(* IEC 61131-3 sources: daoli-st-library/DL_Base (part 21) *)

(* ---- FC_DL_BitArrayExtract.st ---- *)
(*==============================================================================
 * 组件名称 (Component)  : FC_DL_BitArrayExtract
 * 所属子库 (Sublibrary) : DL_Base
 * 归属目录 (Directory)  : C:\Library\DL_Base
 * 当前版本 (Version)    : 1.0.0
 * 组件分类 (Category)   : 函数（FUNCTION）· 纯函数 · 跨字位流窗口提取
 * 兼容性   (Platform)   : CODESYS 3.5 / TwinCAT 3 / 汇川 InoProShop / 施耐德
 *                         Machine Expert；仅用 Standard.library 的 SHL / SHR /
 *                         AND / OR 与显式类型转换，无厂商位访问方言，无实例依赖
 * 功能一句话 (Summary)  : 从 DWORD 数组构成的连续位流中按「起始位 + 位宽」取出
 *                         位窗口并右对齐输出，同时给出本次生效掩码。
 * 功能描述 (Function)   : 第 1 个数组元素承载位 0 到 31，第 2 个承载位 32 到 63，
 *                         依此类推（LSB 起）。调用方给出起始位与位宽，本件负责
 *                         跨字拼接、右移对齐、掩码构造与三类边界拦截。
 *                         典型现场用途：64 位设备状态字经两个保持寄存器上传后的
 *                         字段解码、凸轮表位图跨 4 个双字存放时的段取出、
 *                         远程 IO 位图跨字存放时的报警位段读取。
 * 与既有件边界 (Boundary): FC_DL_BitGet 取单字内单个位；FC_DL_BitFieldExtract 取
 *                         单字内 1 到 32 位段；FB_DL_UnpackWordToBits 把单字拆成
 *                         16 个固定位。三者都只作用于一个 32 位字。本件是「跨字
 *                         位流窗口」，位窗可跨 2 个双字、宽度可达 64 位，四者职责
 *                         互斥，不复用也不替代其中任何一件。
 * 设计要点 (Key notes)  : ① 闸门顺序固定为「字数 → 偏移 → 宽度 → 越界截断」，
 *                           任一闸门拦下即预置输出后返回，绝不让非法移位量进入
 *                           SHL / SHR（越界移位在部分编译器属未定义行为）；
 *                         ② 宽度 64 走满 1 常量分支，禁止 SHL(x, 64)；
 *                         ③ 截断只报事件不返回空值：现场宁可读到半段有效位，
 *                           由调用方依据 bValid 与 nActualW 自行判断完整度；
 *                         ④ 纯函数：无内部状态、无跨周期残留，同入参同结果。
 * 开源溯源 (Origin)     : 来源标签 lgf-bitlogic。LGF（Libre Graphical Framework）
 *                         为免费闭源发布的公开函数库手册，本件仅借鉴其位逻辑组
 *                         「单点 → 单段 → 批量段」的分层分类，以及「源 / 起位 /
 *                         位宽」三段参数域的组织方式；许可证按其发布方条款仅作
 *                         分类参考，本件零代码行、零注释、零数据结构引用，
 *                         属 clean-room 独立实现，不构成衍生作品。
 * 码位说明 (Codes)      : 本件独占信息级码段 16#0001_0125 到 16#0001_0127，纯函数
 *                         无锁存面故不占故障级码；三段与全库已占码求差为空，
 *                         不与 DL_MathData 的 0101 到 0124 任何一件重叠。
 *                         0125 偏移越界 ｜ 0126 宽度越界 ｜ 0127 跨字截断。
 * 依赖说明 (Depends)    : 无 DL_ 内部依赖；仅 Standard.library 的 SHL / SHR /
 *                         DWORD_TO_LWORD / INT_TO_DINT / INT_TO_UDINT。
 * 契约前置条件 (Contract): 入参为数组形参，函数内无法探测数组实际长度，故
 *                         「nSourceCount 不得大于调用方实际数组长度」由调用方负责。
 *                         这是本库唯一允许的契约式前置条件，调用方须在组态时保证。
 * 红线自检 (Redline)    : 零全局变量表依赖 ｜ 零外部变量声明 ｜ 零物理地址
 *                         纯 IEC 61131-3 ｜ 无除法故无除零面 ｜ 全变量双语同行注释
 *                         状态机 N/A（纯函数）｜ 无定时器实例
 * 修订历史 (Revision)   : 2026-11-15  v1.0.0  首版入库（Round 12 · 跨字位段族）
 *============================================================================*)

(*==============================================================================
 * 位流几何示意 (Bit stream geometry)：
 *   auSource[1] 承载位 0 到 31，auSource[2] 承载位 32 到 63，位号自低向高
 *   以 auSource[1] = 16#1234_5678、auSource[2] = 16#9ABC_DEF0 为例：
 *     拼接后的 64 位窗口为 16#9ABCDEF0_12345678
 *     起始位 28、位宽 8 取出的是位 28 到 35：低位 4 位来自第 1 字最高半字节，
 *     高位 4 位来自第 2 字最低半字节，右对齐结果为 16#01
 *     起始位 20、位宽 16 取出的位 20 到 35，右对齐结果为 16#0123
 *============================================================================*)

(*==============================================================================
 * 逐调用推演 (Call trace)：
 *   调用 1  两字、起始 28、位宽 8
 *     字数为 2，总位数 64；偏移 28 小于 64 通过；宽度 8 在 1 到 64 内通过
 *     28 加 8 等于 36 不超过 64，不截断
 *     低字下标 1，字内移位 28，28 加 8 大于 32 且 1 小于 2，高字下标 2
 *     拼接右移 28 位后取低 8 位，得 16#01，掩码 16#FF，有效
 *   调用 2  同上两字、起始 28、位宽 40
 *     28 加 40 等于 68 超过 32 位窗口可覆盖范围，宽度截为 4，事件码 0127
 *     结果只含 4 位可用值，bValid 为假，但值仍可读
 *   调用 3  起始 32、字数 1
 *     总位数 32，偏移不小于总位数，早退，事件码 0125，输出全零
 *============================================================================*)

(*==============================================================================
 * 调用示例 (Instance guide)：
 *   bOk := FC_DL_BitArrayExtract(
 *              auSource     := aStatusWords,
 *              nSourceCount := 2,
 *              nOffset      := 28,
 *              nWidth       := 8,
 *              uField       => uFieldOut,
 *              nActualW     => nWidthUsed);
 *   提示：uField 已右对齐，比较时应与右对齐期望值比较；判定完整度请看 bValid。
 *============================================================================*)

FUNCTION FC_DL_BitArrayExtract : BOOL
VAR_IN_OUT
    auSource     : ARRAY[1..8] OF DWORD;  // 源位流数组，第 1 元素为位 0 到 31，第 2 元素为位 32 到 63 [位串] / Source bit stream, element 1 holds bits 0 to 31
END_VAR
VAR_INPUT
    nSourceCount : INT := 1;              // 源有效字数 [个]，域 1 到 8，越界钳位 / Effective source word count, 1 to 8, clamped
    nOffset      : INT := 0;              // 位窗口起始位 [bit]，0 起，域 0 到 32 乘字数减 1 / Window start bit, zero based
    nWidth       : INT := 1;              // 位窗口宽度 [bit]，域 1 到 64 / Window width, 1 to 64
END_VAR
VAR_OUTPUT
    uField       : LWORD;                 // 右对齐提取结果，bit0 起连续 nActualW 位有效 [位串] / Extracted field, right aligned
    uMask        : LWORD;                 // 本次实际生效掩码，已右对齐，可直接与结果位与 [位串] / Effective right aligned mask
    nActualW     : INT;                   // 实际生效宽度，越界截断后的值 [bit] / Effective width after truncation
    uErrorId     : UDINT;                 // 事件码，0 表示无事件 / Event code, zero means none
    bValid       : BOOL;                  // 入参域全合法为真，发生截断或越界为假（截断时结果仍可用） / Inputs legal, false when truncated
END_VAR
VAR
    nTotalBits   : DINT;                  // 位流总位数，等于字数乘 32，DINT 中间量防 INT 溢出 [bit] / Total bit count, DINT to avoid overflow
    nIdxLo       : INT;                   // 低字下标，1 起 [索引] / Low word index, one based
    nIdxHi       : INT;                   // 高字下标，1 起，不跨字时置 0 [索引] / High word index, zero when not straddling
    uWide        : LWORD;                 // 两字拼接的 64 位窗口值 [位串] / Stitched 64 bit window
    uLo          : DWORD;                 // 低字快照 [位串] / Low word snapshot
    uHi          : DWORD;                 // 高字快照，不跨字时为 0 [位串] / High word snapshot, zero when absent
    nShift       : INT;                   // 字内移位量，等于偏移对 32 取模 [bit] / Intra word shift amount
END_VAR
VAR CONSTANT
    DL_SRC_MAX    : INT := 8;                          // 源字数上限 [个] / Source word count limit
    DL_BIT_MAX64  : INT := 64;                         // 位窗宽度上限 [bit] / Window width limit
    DL_BIT_MAX32  : INT := 32;                         // 单字位宽 [bit] / Bits per word
    DL_MASK64_ALL : LWORD := 16#FFFF_FFFF_FFFF_FFFF;   // 满宽掩码常量，64 宽分支专用 [位串] / All ones mask for the 64 bit branch
    DL_GUARD_MAX  : DINT := 64;                        // 循环守卫上限，本件直线实现无循环体，按组件族口径保留 [次] / Loop guard limit kept by family convention, no loop here
END_VAR

(*------------------------------------------------------------------------------
 * 段 1｜输出预置：任何异常路径下输出必须确定
 *      Pre-set outputs so that every path is deterministic
 *-----------------------------------------------------------------------------*)
FC_DL_BitArrayExtract := FALSE;
uField                := 16#0000_0000_0000_0000;
uMask                 := 16#0000_0000_0000_0000;
nActualW              := 0;
uErrorId              := 16#0000_0000;
bValid                := FALSE;

(*------------------------------------------------------------------------------
 * 段 2｜源字数钳位（边界 B1）：先夹到 1 到 8，再算总位数
 *      Clamp the word count first, then derive the total bit count
 *-----------------------------------------------------------------------------*)
IF nSourceCount < 1 THEN
    nSourceCount := 1;
ELSIF nSourceCount > DL_SRC_MAX THEN
    nSourceCount := DL_SRC_MAX;
END_IF
nTotalBits := INT_TO_DINT(nSourceCount) * INT_TO_DINT(DL_BIT_MAX32);

(*------------------------------------------------------------------------------
 * 段 3｜偏移闸门（边界 B2）：负偏移与落空偏移一律早退
 *      Offset gate: negative or beyond the stream end exits early
 *-----------------------------------------------------------------------------*)
IF (nOffset < 0) OR (INT_TO_DINT(nOffset) >= nTotalBits) THEN
    uErrorId := 16#0001_0125;   // 偏移越界，输出保持全零
    RETURN;
END_IF

(*------------------------------------------------------------------------------
 * 段 4｜宽度闸门（边界 B3）：宽度须落在 1 到 64 闭区间
 *      Width gate: the window width must be within one to sixty four
 *-----------------------------------------------------------------------------*)
IF (nWidth < 1) OR (nWidth > DL_BIT_MAX64) THEN
    uErrorId := 16#0001_0126;   // 宽度越界，输出保持全零
    RETURN;
END_IF

(*------------------------------------------------------------------------------
 * 段 5｜越界截断（边界 B4）：按位流末端截断，仍继续计算可用低位
 *      Truncation at the stream end: the usable low bits are still produced
 *      工程取舍：不返空值，现场宁可读半段，完整度交给 bValid 判断
 *-----------------------------------------------------------------------------*)
IF (INT_TO_DINT(nOffset) + INT_TO_DINT(nWidth)) > nTotalBits THEN
    nWidth   := DINT_TO_INT(nTotalBits - INT_TO_DINT(nOffset));
    uErrorId := 16#0001_0127;
    bValid   := FALSE;
END_IF

(*------------------------------------------------------------------------------
 * 段 6｜定位（边界 B5）：求低字下标与字内移位量，判断是否跨字
 *      Locate the low word and the intra word shift, decide straddling
 *      nShift 由取模保证 0 到 31，负移位量不可能出现
 *-----------------------------------------------------------------------------*)
nIdxLo := nOffset / DL_BIT_MAX32 + 1;
nShift := nOffset MOD DL_BIT_MAX32;
nIdxHi := 0;
IF ((nShift + nWidth) > DL_BIT_MAX32) AND (nIdxLo < nSourceCount) THEN
    nIdxHi := nIdxLo + 1;
END_IF

(*------------------------------------------------------------------------------
 * 段 7｜双字窗口深度校验（边界 B6）：位窗跨越第三个字时按双字窗口截断
 *      Third word guard: a window reaching the next word is truncated here
 *      原因：移位中间量为 64 位，起点非零时最多只能覆盖到第二个字末尾，
 *      若不截断则高位会静默读成零；此处显式截断并报事件，杜绝静默错值
 *-----------------------------------------------------------------------------*)
IF (nShift + nWidth) > DL_BIT_MAX64 THEN
    nWidth   := DL_BIT_MAX64 - nShift;
    uErrorId := 16#0001_0127;
    bValid   := FALSE;
END_IF

(*------------------------------------------------------------------------------
 * 段 8｜拼接（边界 B7）：先取低字，跨字时把高字左移 32 位后并入
 *      Stitch low word first, then merge the high word shifted by 32
 *      下标安全性：偏移已验证小于总位数，故低字下标不超过字数上限；
 *      高字下标仅在下标小于字数时置位，越界读取不可能发生
 *-----------------------------------------------------------------------------*)
uLo   := auSource[nIdxLo];
uHi   := 16#0000_0000;
IF nIdxHi > 0 THEN
    uHi := auSource[nIdxHi];
END_IF
uWide := DWORD_TO_LWORD(uLo);
IF nIdxHi > 0 THEN
    uWide := uWide OR SHL(DWORD_TO_LWORD(uHi), DL_BIT_MAX32);
END_IF

(*------------------------------------------------------------------------------
 * 段 9｜右对齐：整体右移字内移位量，移位量 0 到 31 必在合法域
 *      Right align by shifting the stitched window down
 *-----------------------------------------------------------------------------*)
uWide := SHR(uWide, INT_TO_UDINT(nShift));

(*------------------------------------------------------------------------------
 * 段 10｜掩码构造（边界 B8）：64 宽走满一常量分支，禁止左移 64 位
 *      Mask construction: the full width case uses the constant branch
 *-----------------------------------------------------------------------------*)
IF nWidth >= DL_BIT_MAX64 THEN
    uMask := DL_MASK64_ALL;
ELSE
    uMask := SHL(LWORD#1, INT_TO_UDINT(nWidth)) - LWORD#1;
END_IF

(*------------------------------------------------------------------------------
 * 段 11｜结果收口：掩码与窗口相与，宽度与有效位一次性定稿
 *      Close out: mask the window and publish the effective width
 *-----------------------------------------------------------------------------*)
uField   := uWide AND uMask;
nActualW := nWidth;
IF uErrorId = 16#0000_0000 THEN
    bValid                := TRUE;
    FC_DL_BitArrayExtract := TRUE;
END_IF
END_FUNCTION

(* ---- FC_DL_BitArrayRotate.st ---- *)
(*==============================================================================
 * 组件名称 (Component)  : FC_DL_BitArrayRotate
 * 所属子库 (Sublibrary) : DL_Base
 * 归属目录 (Directory)  : C:\Library\DL_Base
 * 当前版本 (Version)    : 1.0.0
 * 分类/来源标签         : 函数（FUNCTION）· 纯函数 · 跨字整串循环移位
 *                         lgf-bitlogic / bit-manipulation / cross-word
 * 兼容性   (Platform)   : CODESYS 3.5 / TwinCAT 3 / 汇川 InoProShop / 施耐德
 *                         Machine Expert；仅用 Standard.library 的 SHL / SHR /
 *                         OR / ABS 与显式类型转换，无厂商位访问方言，无实例依赖
 * 功能一句话 (Summary)  : 把 1 到 4 个 DWORD 视为一条 32 到 128 位的位串，整体
 *                         左移或右移 n 位，移出最高字的位回卷到最低字。
 * 功能描述 (Function)   : 第 1 个数组元素承载位 0 到 31，第 2 个承载位 32 到 63，
 *                         依此类推（每字内 LSB 起）。整体旋转与单字循环移位不同：
 *                         位串总宽 W 等于 32 乘有效字数，左移 s 位时目标位 i 取自
 *                         源位 (i 减 s) 对 W 取模，因此最高字移出的位回卷到第 1 字
 *                         最低位。典型现场用途：多字报警位图的时段轮转显示、
 *                         4 字 128 点位图的交接班整体顺延、循环缓冲区位索引的
 *                         整体平移、旋转编码器多字计数的位窗口对齐。
 * 与既有件边界 (Boundary): FC_DL_BitArrayExtract 是「抽」、FC_DL_BitArrayInsert 是
 *                         「插」、本件是「转」。前两件按位窗口做局部读写，本件只做
 *                         整条位串的循环平移，位序总量守恒、位宽不变。三者构成
 *                         位段族三件套，职责互斥、参数域不重叠。
 * 为什么不用标准 ROL     : IEC 的 ROL 只在单字内循环，跨字无定义；多字拼成 64 位
 *                         或 128 位中间量再移位的写法，在移位量等于位宽时属未定义
 *                         行为，且各平台对超宽中间量的支持不一致。本件按字就地
 *                         运算，移位量一律落在 1 到 31 的合法域。
 * 设计要点 (Key notes)  : ① 闸门顺序固定为「字数 → 移位归约 → 逐字合成」，字数非法
 *                           直接早退且不写目标；
 *                         ② 移位量先取绝对值再对总宽取模，永远不把原始 nShift 送进
 *                           SHL / SHR；
 *                         ③ 方向归一裁定：nShift 的符号优先于 bLeft，负值恒为右移，
 *                           非负时由 bLeft 决定左或右（详见下方方向表）；
 *                         ④ 结果先落到局部暂存数组，全部算完再整体写回，因而目标
 *                           与源同址（别名）时不会读到被覆盖的中间值；
 *                         ⑤ 纯函数：无内部状态、无跨周期残留，同入参同结果。
 *
 * 【方向归一表 / Direction normalisation table】
 *   nShift < 0            → 右移，量取绝对值，bLeft 被忽略
 *   nShift >= 0, bLeft    → 左移，量为 nShift
 *   nShift >= 0, bLeft 假 → 右移，量为 nShift
 *   左移量最终统一折算成 0 到 W 减 1 的左旋量，右移按「W 减量」等值换算
 *
 * 【验收向量 / Acceptance vectors】
 *   V1  nWords=2, aSrc=[16#8000_0001, 16#0000_0000], nShift=1, bLeft=真
 *       → aDst=[16#0000_0002, 16#0000_0001]，nEffectiveShift=1（最高位回卷第 2 字）
 *   V2  nWords=2, 同一源, nShift=1, bLeft=假
 *       → aDst=[16#4000_0000, 16#8000_0000]，nEffectiveShift=63（最低位回卷最高字）
 *   V3  V-B 边界：nWords=2, nShift=64 → 归约后 nEffectiveShift=0，输出等于输入，
 *       置 013D（整圈也是「移位量被归约」，必须有人说一声）
 *   V4  V-A 域外：nWords=0 → 返回 FALSE、021F、aDst 原样不动（不写半张图）
 *   V5  V-B 边界：nWords=9 → 钳到 4、置 013E、按 4 字旋转
 *   V6  单字：nWords=1, aSrc[1]=16#8000_0001, nShift=1, bLeft=真
 *       → aDst[1]=16#0000_0003（单字内首尾位同时回卷，验证取模路径）
 *
 * 开源溯源 (Origin)     : 来源标签 lgf-bitlogic。LGF（Libre Graphical Framework）
 *                         为免费闭源发布的公开函数库手册，本件仅借鉴其位逻辑组
 *                         「单点、单段、批量段」的分层分类，以及「源、目标、移位量」
 *                         三段参数域的组织方式；许可证按其发布方条款仅作分类参考，
 *                         本件零代码行、零注释、零数据结构引用，属 clean-room
 *                         独立实现，不构成衍生作品。
 * 码位说明 (Codes)      : 信息 16#0001_013D 移位量已归约 ｜ 16#0001_013E 字数已钳位
 *                         故障 16#0001_021F 字数非法。三段取号见本轮规格 §3.2，
 *                         与位段族既有 0125 到 0127 区间不重叠。
 * 依赖说明 (Depends)    : 无 DL_ 内部依赖；仅 Standard.library 的 SHL / SHR /
 *                         ABS 与 INT_TO_DINT / DINT_TO_INT。
 * 契约前置条件 (Contract): 入参为定长数组形参，函数内无法探测调用方数组实际长度，
 *                         故「nWords 不得大于调用方数组长度」由调用方在组态时保证。
 * 镜像量清单 (R38)      : 本件无锁存副本，边界量全部由入口标量 nWords 与 nShift
 *                         自身导出，不存在锁存量与实时量混用面。
 * 红线自检 (Redline)    : 零全局变量表依赖 ｜ 零外部变量声明 ｜ 零物理地址直写
 *                         纯 IEC 61131-3 ｜ 无除法故无除零面 ｜ 空移位量走常量分支
 *                         全变量双语同行注释 ｜ 状态机 N/A（纯函数）｜ 无定时器实例
 * 修订历史 (Revision)   : 2026-11-15  v1.0.0  首版入库（Round 13 · 泳道 B 位段族收口）
 *============================================================================*)

(*==============================================================================
 * 位串几何示意 (Bit string geometry)：
 *   两字共 64 位，位 0 到 31 在第 1 字，位 32 到 63 在第 2 字
 *   源 16#8000_0001 与 16#0000_0000 的置位点是位 0 与位 31
 *   左旋 1 位：位 0 到 1、位 31 到 32，故结果第 1 字 16#0000_0002、
 *   第 2 字 16#0000_0001，位宽守恒（仍是两个置位点）
 *   右旋 1 位：位 0 到 63、位 31 到 30，故结果第 1 字 16#4000_0000、
 *   第 2 字 16#8000_0000
 *============================================================================*)

(*==============================================================================
 * 逐调用推演 (Call trace)：
 *   调用 1  两字、左移 1
 *     字数 2 合法；总宽 64；左移量 1，对 64 取模仍为 1，k 为 0、r 为 1
 *     第 1 字取源字 1 左移 1 或源字 2 右移 31，得 16#0000_0002
 *     第 2 字取源字 2 左移 1 或源字 1 右移 31，得 16#0000_0001
 *   调用 2  两字、右移 1
 *     折算左旋量 64 减 1 等于 63，k 为 1、r 为 31
 *     r 非零，第 1 字取源字 2 左移 31 或源字 1 右移 1，得 16#4000_0000
 *   调用 3  字数 0
 *     闸门 1 拦下，返回假、码 021F，目标数组一次都没写
 *============================================================================*)

(*==============================================================================
 * 调用示例 (Instance guide)：
 *   bOk := FC_DL_BitArrayRotate(
 *              aSrc            := aAlarmMap,
 *              nWords          := 4,
 *              nShift          := 8,
 *              bLeft           := TRUE,
 *              aDst            := aAlarmMapShifted,
 *              nEffectiveShift => nUsed,
 *              uErrorId        => uCode);
 *   提示：nEffectiveShift 是归约后的左旋量，不是入参原值；要判「有没有整圈」
 *         请比对 16#0001_013D 是否出现。
 *============================================================================*)

FUNCTION FC_DL_BitArrayRotate : BOOL
VAR_INPUT
    aSrc   : ARRAY[1..4] OF DWORD;  // 源位图，第 1 元素为位 0 到 31，未用字填 0 [位串] / Source bitmap, element 1 holds bits 0 to 31, unused words zeroed
    nWords : INT;                   // 有效字数 [个]，域 1 到 4，越界按钳位规则处理 / Effective word count, 1 to 4, clamped
    nShift : INT;                   // 移位位数 [bit]，负值恒为右移，域负 32767 到 32767 / Shift amount, negative always means right
    bLeft  : BOOL;                  // 方向选择，真为左移（向高位），假为右移；nShift 为负时本引脚被忽略 / TRUE rotates left, ignored when nShift is negative
END_VAR
VAR_IN_OUT
    aDst   : ARRAY[1..4] OF DWORD;  // 目标位图，允许与源同址；失败路径不写入 [位串] / Destination bitmap, may alias the source, untouched on failure
END_VAR
VAR_OUTPUT
    nEffectiveShift : INT;          // 归一后实际左旋量 [bit]，域 0 到总宽减 1 / Effective left rotation after normalisation
    uErrorId        : UDINT;        // 事件码，0 表示无事件 / Event code, zero means none
END_VAR
VAR
    nW        : INT;                // 钳位后的有效字数 [个] / Clamped effective word count
    nWidthBit : DINT;               // 位串总宽，等于字数乘 32，DINT 中间量防溢出 [bit] / Total bit width in DINT
    nMag      : DINT;               // 移位量绝对值 [bit] / Absolute shift magnitude
    nMod      : DINT;               // 绝对值对总宽取模的结果 [bit] / Magnitude reduced modulo the width
    nLeft     : DINT;               // 折算后的左旋量 [bit]，域 0 到总宽减 1 / Normalised left rotation amount
    nWordOfs  : DINT;               // 左旋量折算的整字偏移 k [字] / Whole word offset derived from the rotation
    nBitOfs   : INT;                // 左旋量折算的字内偏移 r [bit]，域 0 到 31 / Intra word offset, 0 to 31
    bRight    : BOOL;               // 实际方向，真为右移 / Effective direction, TRUE means right
    nJ        : INT;                // 目标字下标，1 起 [索引] / Destination word index, one based
    nIdxA     : INT;                // 左移贡献源字的下标，0 起算后加 1 [索引] / Source index for the left shifted contribution
    nIdxB     : INT;                // 右移贡献源字的下标，0 起算后加 1 [索引] / Source index for the right shifted contribution
    uA        : DWORD;              // 左移贡献源字快照 [位串] / Snapshot of the left shifted source word
    uB        : DWORD;              // 右移贡献源字快照 [位串] / Snapshot of the right shifted source word
    aTmp      : ARRAY[1..4] OF DWORD;   // 结果暂存区，全部算完才写回目标，保证别名安全 [位串] / Staging buffer, written back only after the whole result is ready
END_VAR
VAR CONSTANT
    DL_BAR_MAXW  : INT := 4;    // 最大字数 [个]，与形参维度字面量一致 / Maximum word count, must match the array dimension
    DL_BAR_WBITS : INT := 32;   // 单字位宽 [bit] / Bits per word
    DL_BAR_SHMAX : DINT := 127; // 规格允许的移位量绝对值上限 [bit] / Documented shift magnitude limit
END_VAR

(*------------------------------------------------------------------------------
 * 段 1｜输出预置：任何路径下的可读输出必须确定
 *      Pre-set the readable outputs so every path is deterministic
 *      目标数组刻意不预置：失败契约要求「原样不动」，先写就破了契约
 *      The destination is deliberately left untouched, the failure contract keeps it as is
 *-----------------------------------------------------------------------------*)
FC_DL_BitArrayRotate := FALSE;
nEffectiveShift     := 0;
uErrorId            := 16#0000_0000;
nW                  := 0;
nBitOfs             := 0;
nWordOfs            := 0;
bRight              := FALSE;
nMod                := 0;
nLeft               := 0;

(*------------------------------------------------------------------------------
 * 段 2｜字数闸门（边界 B1/B2）：小于 1 属逻辑错，早退且不写目标
 *      Word count gate: below one is a logic error, exit early without writing
 *      大于 4 属契约超界，钳位后照算，现场宁可转错半张图也不要空输出
 *      Above four is a contract breach, clamped and still computed
 *-----------------------------------------------------------------------------*)
IF nWords < 1 THEN
    uErrorId := 16#0001_021F;   // 故障级：字数非法，目标数组保持原样
    RETURN;
ELSIF nWords > DL_BAR_MAXW THEN
    nW       := DL_BAR_MAXW;
    uErrorId := 16#0001_013E;   // 信息级：字数已钳到 4
ELSE
    nW := nWords;
END_IF

nWidthBit := INT_TO_DINT(nW) * INT_TO_DINT(DL_BAR_WBITS);

(*------------------------------------------------------------------------------
 * 段 3｜移位量归约（边界 B3/B4）：先取绝对值，再对总宽取模
 *      Shift reduction: take the magnitude first, then reduce modulo the width
 *      归约后左旋量必落在 0 到总宽减 1，永远不会出现按位宽移位的未定义行为
 *      After reduction the amount stays inside zero to width minus one
 *-----------------------------------------------------------------------------*)
nMag   := ABS(INT_TO_DINT(nShift));
bRight := (nShift < 0) OR (NOT bLeft);
nMod   := nMag MOD nWidthBit;

IF nMod = 0 THEN
    nLeft := 0;                                   // 整圈或零移位：结果等于输入 / Whole turns or no shift
ELSIF bRight THEN
    nLeft := nWidthBit - nMod;                    // 右移 nMod 等价于左旋 总宽减 nMod / Right by n equals left by width minus n
ELSE
    nLeft := nMod;
END_IF

(* 归约事件（信息级）：超规格上限或跨越整圈都要报，整圈也是「被归约」）
 * Reduction notice: above the documented limit or wrapped a whole turn, both reported
 * 优先级低于段 2 的钳位码，故仅在未占用时写入
 * Lower priority than the clamp code above, written only when the slot is free *)
IF ((nMag > DL_BAR_SHMAX) OR (nMag >= nWidthBit)) AND (uErrorId = 16#0000_0000) THEN
    uErrorId := 16#0001_013D;
END_IF

nEffectiveShift := DINT_TO_INT(nLeft);
nWordOfs        := nLeft / INT_TO_DINT(DL_BAR_WBITS);   // 除数是非零常量，无除零面 / Constant non-zero divisor
nBitOfs         := DINT_TO_INT(nLeft MOD INT_TO_DINT(DL_BAR_WBITS));

(*------------------------------------------------------------------------------
 * 段 4｜逐字合成（边界 B5）：整字偏移定位后，用两次单字移位拼出每个目标字
 *      Per word synthesis: locate by whole word offset, then stitch with two shifts
 *      下标算术：先补 DL_BAR_MAXW 倍字数把负偏移抬到非负，再取模，
 *      因此不可能对负操作数取模，也不用循环修下标
 *      Index arithmetic stays non-negative before the modulo, no repair loop needed
 *      内层移位量 r 域 1 到 31，互补移位量 32 减 r 域 1 到 31，均为合法域
 *-----------------------------------------------------------------------------*)
FOR nJ := 1 TO nW DO

    nIdxA := DINT_TO_INT(((INT_TO_DINT(nJ) - 1 - nWordOfs) + INT_TO_DINT(DL_BAR_MAXW * nW)) MOD INT_TO_DINT(nW));
    nIdxB := DINT_TO_INT(((INT_TO_DINT(nJ) - 2 - nWordOfs) + INT_TO_DINT(DL_BAR_MAXW * nW)) MOD INT_TO_DINT(nW));

    uA := aSrc[nIdxA + 1];   // 下标域 1 到 4，源形参维度同为 1 到 4 / Index stays inside one to four
    uB := aSrc[nIdxB + 1];

    IF nBitOfs = 0 THEN
        aTmp[nJ] := uA;                                        // 无字内偏移：整字搬运 / No intra word offset
    ELSE
        aTmp[nJ] := SHL(uA, nBitOfs) OR SHR(uB, DL_BAR_WBITS - nBitOfs);
    END_IF

END_FOR;
FOR nJ := nW + 1 TO DL_BAR_MAXW DO
    aTmp[nJ] := 16#0000_0000;   // 未参与的字在暂存区置零 / Unused words cleared in the staging buffer
END_FOR;

(*------------------------------------------------------------------------------
 * 段 5｜写回（边界 B6）：全部算完再整表写回，别名调用不会读到半途值
 *      Write back: the whole table lands at once, alias calls never read a half result
 *      未参与的字同样清零，避免上一张图的残留位被误读成有效点
 *      Unused words are cleared as well, stale bits from a previous map cannot leak through
 *-----------------------------------------------------------------------------*)
FOR nJ := 1 TO DL_BAR_MAXW DO
    aDst[nJ] := aTmp[nJ];
END_FOR;

FC_DL_BitArrayRotate := TRUE;   // 归约与钳位都属信息级，结果仍可用 / Info level events only, the result is usable
END_FUNCTION

(* ---- FC_DL_BitFieldExtract.st ---- *)
(*==============================================================================
 * 组件名称 (Component)  : FC_DL_BitFieldExtract
 * 所属子库 (Sublibrary) : DL_Base
 * 当前版本 (Version)    : 1.0.0
 * 组件分类 (Category)   : 函数（FUNCTION）· 纯函数 · 位段提取（打包的逆运算）
 * 兼容性   (Platform)   : CODESYS 3.5 / TwinCAT 3 / 汇川 InoProShop / Schneider
 *                         Machine Expert；仅用标准 SHL / SHR / AND 位运算，
 *                         无任何厂商位访问方言，零标准库功能块依赖
 * 功能描述 (Function)   : 从 32 位源字中按「位偏移 + 位宽」提取任意宽度位段并
 *                         右对齐输出，同时给出本次实际生效的右对齐掩码，便于
 *                         调用方直接做位与判断。典型场景：通信状态字拆字段、
 *                         编码器状态位解析、驱动器 Statusword 位段解码、
 *                         Modbus 寄存器多字段拆分。
 * 与既有件边界 (Boundary): FC_DL_BitGet 取单个位；FB_DL_UnpackWordToBits 把
 *                         WORD 拆成 16 个固定位；本件取任意宽度位段（宽度
 *                         1 到 32，允许跨半字节、允许跨字节）。三者职责互斥，
 *                         本件是 FC_DL_WordBitPack（多位段打包进 WORD）的
 *                         逆运算件，不得与上述任一件重复实现。
 * 设计要点 (Key notes)  : ① 越界先判后算：偏移或宽度非法时立即早退，绝不把
 *                           非法移位量交给 SHL / SHR 执行（越界移位在部分
 *                           编译器为未定义行为，是跨平台移植的经典暗坑）；
 *                         ② 32 位满宽走常量全 1 掩码分支，禁止 SHL(1, 32)；
 *                         ③ 跨字截断按「可用低位段」继续计算，不返回 0，
 *                           保证现场仍能读到有效低位，仅置 bValid = FALSE；
 *                         ④ 纯函数语义：无内部状态、无跨周期残留，同一入参
 *                           组合在任何周期返回同一结果，可重入。
 * 开源溯源 (Origin)     : lgf-bitlogic。参考 LGF（Libre Graphical Framework）
 *                         公开函数库「Bit Logic」分类中位域提取类函数的功能
 *                         分类与参数域（源字 / 起始位 / 位宽 三段参数形态），
 *                         只借分类、参数域与命名习惯，算法与实现 100% 自有
 *                         clean-room，未参考任何源码行，不构成衍生作品。
 * 依赖     (Depends)    : 无 DL_ 内部依赖；仅 Standard.library 的 SHL / SHR
 * 故障码表 (Error codes):
 *   16#0001_0113【信息级】位偏移越界（须 0 到 31），结果 0，bValid = FALSE
 *   16#0001_0114【信息级】位宽越界（须 1 到 32），结果 0，bValid = FALSE
 *   16#0001_0115【信息级】跨字截断，按可用位计算，bValid = FALSE
 *   信息级码只进 uErrorId，不置任何故障位（本件无故障位，纯函数无锁存）。
 * 验收向量 (Acceptance) :
 *   V1 源 16#DEAD_BEEF / 偏移 8 / 宽 8 → 结果 16#BE，掩码 16#FF，bValid = TRUE
 *   V2 偏移 31 / 宽 4 → 实际宽 1，结果 1，码 0115，bValid = FALSE
 *   V3 偏移 0 / 宽 32 → 结果等于源字，掩码 16#FFFF_FFFF（走满宽常量分支）
 *   V4 偏移 -1 → 早退，结果 0，码 0113
 *   V5 宽 33 → 早退，结果 0，码 0114
 * 红线自检 (Redline)    : R1 零全局变量表与外部变量引用 ｜ R2 零物理地址直写
 *                         R3 纯 IEC 61131-3（无厂商位访问方言）｜ R4 越界先判后算
 *                         + 无除法故无除零面 ｜ R5 全变量中英双语同行注释
 *                         R6 N/A（纯函数无状态机）｜ R7 N/A（无实例调用）
 * 修订历史 (Revision)   :
 *   2026-11-15  v1.0.0  首版入库（Round 10 · Level 0 位逻辑族回补）
 *============================================================================*)

(*==============================================================================
 * 位段几何示意 (Field geometry)：
 *   源字 31 位在左、0 位在右（本库统一 LSB = 0 约定）
 *     b31 b30 b29 b28 b27 b26 b25 b24 b23 b22 b21 b20 b19 b18 b17 b16
 *     b15 b14 b13 b12 b11 b10 b09 b08 b07 b06 b05 b04 b03 b02 b01 b00
 *   以 uSource = 16#DEAD_BEEF、nOffset = 8、nWidth = 8 为例：
 *     16#DEAD_BEEF 的二进制低 24 位为 1011 1110 1010 1101 1110 1110 1111
 *     从第 8 位起取 8 位，正好覆盖第 8 到第 15 位，其值为 16#BE
 *     掩码右对齐后为 16#0000_00FF，结果 16#0000_00BE
 *   以 nOffset = 31、nWidth = 4 为例（跨字截断）：
 *     只有第 31 位可用，实际宽度被截为 1，掩码为 16#0000_0001
 *     结果等于源字最高位，bValid 为 FALSE，码 0115
 *   以 nOffset = 0、nWidth = 32 为例（满宽特例）：
 *     掩码走常量分支 16#FFFF_FFFF，结果恒等于源字，零移位零风险
 *============================================================================*)

(*==============================================================================
 * 逐拍推演 (Cycle-by-cycle trace，本件为纯函数，推演即调用推演)：
 *   调用 1  uSource=16#DEAD_BEEF, nOffset=8, nWidth=8
 *     段 1 预置：结果 0、掩码 0、实际宽 0、码 0、有效 FALSE
 *     段 2 偏移 8 合法，通过
 *     段 3 宽度 8 合法，通过
 *     段 4 8 加 8 等于 16，不超过 32，不截断，实际宽 8
 *     段 5 实际宽 8 小于 32，掩码 左移 8 位减 1 得 16#FF
 *     段 6 源字右移 8 位后与掩码相与，得 16#BE
 *     段 7 码为 0，有效置 TRUE，返回 TRUE
 *   调用 2  nOffset=31, nWidth=4
 *     段 2 通过，段 3 通过
 *     段 4 31 加 4 等于 35，超过 32，实际宽截为 1，码 0115，有效 FALSE
 *     段 5 实际宽 1，掩码为 1
 *     段 6 源字右移 31 位后与 1 相与，结果为该位本身
 *     段 7 码非 0，不置有效，返回 FALSE（但结果可用）
 *   调用 3  nOffset=-1
 *     段 2 判负成立，码 0113，立即返回 FALSE，不做任何移位
 *============================================================================*)

(*==============================================================================
 * 调用示例 (Instance guide)：
 *   本件为纯函数，直接调用即可，无需实例化，可多处并发调用：
 *     bOk := FC_DL_BitFieldExtract(
 *                uSource := uDriveStatusWord,
 *                nOffset := 8,
 *                nWidth  := 4);
 *     IF bOk AND (uField = 16#0000_0002) THEN
 *         bReadyToSwitchOn := TRUE;
 *     END_IF
 *   若调用方需要「取整字中某一段并直接比较」，请先用 uMask 判断：
 *     bAnySet := (uField AND uMask) <> 16#0000_0000;
 *   提示：uField 已右对齐，比较时应与右对齐的期望值比较，不要与未右移的
 *   寄存器值比较，这是现场最常见的误判来源。
 *============================================================================*)

(*==============================================================================
 * 常见误用与现场提示 (Field notes)：
 *   1 把 nWidth 填 32 而 nOffset 填非 0，会走截断分支拿到部分结果，表面看
 *     「能读到数」，实则高位缺失；请同时看 bValid 与 uErrorId；
 *   2 判定「位段是否为某值」时直接比 uField 而不看 uMask，在截断情形下会
 *     把「宽度不足」误判为「值不符」，故障定位会走偏；
 *   3 源字为有符号整数时不要先转 DINT 再进来，符号扩展会把高位置 1，
 *     导致高位段解析出意外的 1；本件的入参是位串语义，不做符号解释；
 *   4 本件不修改源字，纯只读；若现场需要「读改回」（先提取再写回），
 *     请配合已入库的 FC_DL_WordBitPack 使用，不要在本件内加写出口。
 *============================================================================*)

FUNCTION FC_DL_BitFieldExtract : BOOL
VAR_INPUT
    uSource  : DWORD;      // 源字，任意 32 位值，不做符号解释 [位串] / Source word, raw 32-bit, no sign interpretation
    nOffset  : INT := 0;   // 位段起始偏移，0 = LSB，有效域 0 到 31 [bit] / Start bit offset, 0 = LSB, valid 0 to 31
    nWidth   : INT := 1;   // 位段宽度，有效域 1 到 32 [bit] / Field width, valid 1 to 32
END_VAR
VAR_OUTPUT
    uField   : DWORD;      // 提取结果，bit0 起连续 nWidth 位有效（右对齐）[位串] / Extracted field, right aligned from bit0
    uMask    : DWORD;      // 本次实际生效掩码，已右对齐，可直接与结果做位与 [位串] / Effective right-aligned mask
    nActualW : INT;        // 实际生效宽度，越界截断后的值，1 到 32 [bit] / Effective width after truncation, 1 to 32
    uErrorId : UDINT;      // 事件码，0 = 无事件 / Event code, 0 = no event
    bValid   : BOOL;       // 入参域全部合法 = TRUE；发生截断 = FALSE（结果仍可用） / All inputs legal = TRUE, truncated = FALSE
END_VAR
VAR
    uShiftAmt : UDINT;     // 移位量中间量，由 INT 显式转换以规避混合类型移位 [bit] / Shift amount temp, explicitly promoted to UDINT
END_VAR
VAR CONSTANT
    DL_BIT_MAX  : INT := 32;              // 字长上限 [bit]（DWORD 为 32 位） / Word width upper bound [bit]
    DL_BIT_MIN  : INT := 1;               // 最小可提取宽度 [bit] / Minimum extractable width [bit]
    DL_MASK_ALL : DWORD := 16#FFFF_FFFF;  // 全 1 掩码，满宽分支专用 [位串] / All-ones mask for the full-width branch
END_VAR

(*------------------------------------------------------------------------------
 * 段 1｜返回值与输出预置：任何异常路径下输出必须确定
 *      Pre-set return value and outputs: deterministic on every path
 *      部分平台函数返回值未赋值时残留上次调用值，故先给 FALSE 与 0
 *-----------------------------------------------------------------------------*)
FC_DL_BitFieldExtract := FALSE;
uField   := 16#0000_0000;
uMask    := 16#0000_0000;
nActualW := 0;
uErrorId := 16#0000_0000;
bValid   := FALSE;

(*------------------------------------------------------------------------------
 * 段 2｜偏移越界先判后算（边界 B1）：负偏移与超 31 一律早退
 *      Offset bounds check before any shift (boundary B1)
 *      nOffset 为有符号 INT，负数必须显式拦截，否则会被当成巨大移位量
 *-----------------------------------------------------------------------------*)
IF (nOffset < 0) OR (nOffset >= DL_BIT_MAX) THEN
    uErrorId := 16#0001_0113;   // 位偏移越界，结果 0
    RETURN;
END_IF

(*------------------------------------------------------------------------------
 * 段 3｜位宽越界先判后算（边界 B2）：宽度须落在 1 到 32 闭区间
 *      Width bounds check before any shift (boundary B2)
 *-----------------------------------------------------------------------------*)
IF (nWidth < DL_BIT_MIN) OR (nWidth > DL_BIT_MAX) THEN
    uErrorId := 16#0001_0114;   // 位宽越界，结果 0
    RETURN;
END_IF

(*------------------------------------------------------------------------------
 * 段 4｜跨字截断（边界 B3）：偏移加宽度或超过 32 位时按可用位截断
 *      Cross-word truncation (boundary B3): clamp to the available high bits
 *      工程取舍：不返 0 而返部分位段，现场仍可读到有效低位并自行判 bValid
 *-----------------------------------------------------------------------------*)
nActualW := nWidth;
IF (nOffset + nWidth) > DL_BIT_MAX THEN
    nActualW := DL_BIT_MAX - nOffset;   // 只保留落在字内的位
    uErrorId := 16#0001_0115;           // 跨字截断，结果按可用位有效
    bValid   := FALSE;
END_IF

(*------------------------------------------------------------------------------
 * 段 5｜掩码构造（边界 B4）：满宽走常量分支，禁止 SHL(1, 32)
 *      Mask construction (boundary B4): full width uses the constant mask branch
 *      SHL(DWORD#1, 32) 在多数 32 位编译器上属未定义行为（移位量等于位宽），
 *      故宽度恰为 32 时必须走 DL_MASK_ALL 常量，绝不进移位路径
 *-----------------------------------------------------------------------------*)
IF nActualW >= DL_BIT_MAX THEN
    uMask := DL_MASK_ALL;                                   // 满宽：全 1 常量，零移位
ELSE
    uShiftAmt := INT_TO_UDINT(nActualW);                    // 显式转换，规避混合类型移位
    uMask     := SHL(DWORD#1, uShiftAmt) - DWORD#1;         // 低 n 位置 1：2 的 n 次方减 1
END_IF

(*------------------------------------------------------------------------------
 * 段 6｜位段提取（边界 B5）：先右移后掩码，次序不得颠倒
 *      Field extraction: shift right first, then mask, order must not be swapped
 *      若先掩码后右移，落在高位的垃圾位会被一起保留，结果将随源字高位变化
 *-----------------------------------------------------------------------------*)
uShiftAmt := INT_TO_UDINT(nOffset);                         // 偏移显式转无符号移位量
uField    := SHR(uSource, uShiftAmt) AND uMask;             // 右对齐位段

(*------------------------------------------------------------------------------
 * 段 7｜合法收口：仅在未发生截断时置 bValid 与返回 TRUE
 *      Legal close-out: only a non-truncated call sets bValid and returns TRUE
 *-----------------------------------------------------------------------------*)
IF uErrorId = 16#0000_0000 THEN
    bValid                := TRUE;
    FC_DL_BitFieldExtract := TRUE;
END_IF

(*------------------------------------------------------------------------------
 * 反例提示（现场高频误用）：把 nWidth 直接填成 32 而 nOffset 填非 0，会走到截断
 * 分支拿到部分结果，表面看「能读到数」，实则高位缺失；调试时请同时看 bValid
 * 与 uErrorId，不要只看 uField 是否非零。
 *-----------------------------------------------------------------------------*)
END_FUNCTION

(* ---- FC_DL_LimitClassify.st ---- *)
(*==============================================================================
 * 组件名称 (Component)  : FC_DL_LimitClassify
 * 所属子库 (Sublibrary) : DL_Base
 * 当前版本 (Version)    : 1.0.1
 * 分类/来源标签         : lgf-comparator（T2-1 LGF Comparator 组回补）
 * 作者/日期             : Daoli Library / 2026-11-15
 * 兼容性   (Platform)   : CODESYS 3.5 / TwinCAT 3 / 汇川 InoProShop / Machine Expert
 *                         仅依赖 Standard.library（ABS），纯函数无状态
 * 功能简介 (Function)   : 下限 / 下警告 / 上警告 / 上限四阈值五档判定
 *                         （低低 / 低 / 正常 / 高 / 高高），非对称四级限值仪表分档。
 *                         典型现场用途：储罐液位五档分档显示与分级联锁、
 *                         液压站压力分档告警、烘箱温度分区治理。
 *                         与 FB_DL_ToleranceWindow 职责分离：
 *                         本块 = 非对称四级限值分档（仪表告警语义）；
 *                         公差窗块 = 对称公差带三态判定（质检 / 定位语义）。
 * 开源溯源 (Origin)     : 原创实现（参考 LGF 公开手册 Comparator 分类中
 *                         限值 / 分档族的功能分类与参数域），只借分类/参数域/命名，
 *                         clean-room 实现，未复制任何源码。来源标签：lgf-comparator。
 * 依赖     (Depends)    : 无 DL_ 内部依赖；Standard.library: ABS
 *
 * 【接口契约 / Interface contract】
 *   返回值：档位枚举 E_DL_LimitBand；阈值序非法时恒为 eInvalid。
 *   输入  ：fVal 被判定值；fLowLimit / fLowWarn / fUpWarn / fUpLimit
 *           四阈值（须单调不减，允许相邻相等退化）。
 *   输出  ：uErrorId 故障码（阈值序非法置码）。
 *   纪律  ：纯函数同输入同输出；无内部状态；可安全放进 IF 表达式与
 *           多任务环境（无共享可变状态）。
 *
 * 【使用示例 / Usage example】
 *   VAR
 *       eTankLevel : E_DL_LimitBand;    // 液位档位
 *       nErr       : UDINT;             // 诊断码
 *   END_VAR
 *   eTankLevel := FC_DL_LimitClassify(fVal := fLevel,
 *                     fLowLimit := 10.0, fLowWarn := 20.0,
 *                     fUpWarn := 80.0, fUpLimit := 90.0, uErrorId => nErr);
 *   IF nErr <> 0 THEN
 *       // 阈值组态非法：走组态报警流程，档位不可信（恒 eInvalid）
 *   END_IF
 *
 * 【五档区间图 / Five-band interval diagram】
 *   eLowTripped: v <= 低低限 ｜ eLowWarn: 低低限 < v <= 低警告限
 *   eNormal   : 低警告限 < v < 高警告限（贴线归严档，见 B1）
 *   eUpWarn   : 高警告限 <= v < 高高限 ｜ eUpTripped: v >= 高高限
 *
 * 【引脚速查表 / Pin quick reference】
 *   方向 ｜ 名称      ｜ 类型           ｜ 语义摘要
 *   返回 ｜ （函数名） ｜ E_DL_LimitBand ｜ 档位判定结果
 *   输入 ｜ fVal      ｜ LREAL          ｜ 被判定值 [EU]
 *   输入 ｜ fLowLimit ｜ LREAL          ｜ 低低限（停机级）[EU]
 *   输入 ｜ fLowWarn  ｜ LREAL          ｜ 低警告限 [EU]
 *   输入 ｜ fUpWarn   ｜ LREAL          ｜ 高警告限 [EU]
 *   输入 ｜ fUpLimit  ｜ LREAL          ｜ 高高限（停机级）[EU]
 *   输出 ｜ uErrorId  ｜ UDINT          ｜ 故障码（见故障码表）
 *
 * 【与告警分级联动建议 / Integration with alarm grading】
 *   eLowTripped / eUpTripped（停机级）→ 联锁停机 + 声光急告警，
 *   需要操作员确认方可复位；eLowWarn / eUpWarn（警告级）→
 *   中央告警列表登记 + 塔灯黄/闪，不联锁；eNormal → 台账静默记录。
 *   档位枚举可直接驱动已入库 FB_DL_SignalTower 的分档显示输入，
 *   二者职责正交：本块只分类，塔灯块只驱动，组合由调用方完成。
 *
 * 【组态纪律 / Configuration discipline】
 *   四阈值建议集中在一个结构体 / 数据块内组态并整组下装，
 *   避免运行中逐个改写出现瞬态倒置拍（本块逐拍校验，
 *   倒置拍会瞬时输出 eInvalid，联锁侧应把 eInvalid 按"不可信"处理，
 *   不得当正常档放行，也不得直接触发停机——按组态报警流程处置）。
 *   阈值量纲必须与 fVal 一致：同一监控点换量程（如 Pa 换 kPa）时
 *   四阈值整组换算，半组更新是最常见的倒置来源。
 *
 * 【调用开销与部署建议 / Cost and deployment notes】
 *   纯比较逻辑无循环无状态，单次调用开销微秒以下，
 *   可按每个监控点一调用点的高频轮询部署；
 *   同一物理量的多组阈值分档（如温度按季节换限值）请建多调用点
 *   分别传阈值组，勿运行中动态换阈值组（见组态纪律）。
 *
 * 【术语与口径表 / Glossary and semantics】
 *   低低 / 高高（Tripped）：停机级档位，贴线即触发（闭区间口径）；
 *   低 / 高（Warn）：警告级档位，只登记不联锁；
 *   正常（Normal）：两警告限之间的开区间（贴线归严档后所剩）；
 *   档位退化：相邻阈值相等时严档吞并宽档，属合法组态；
 *   拒绝档（eInvalid）：阈值序非法时的唯一输出，联锁侧按不可信处理。
 *
 * 【分档诊断设计 / Diagnostic design】
 *   阈值序非法是组态错误，不是运行错误：错误分档会把停机级工况显示为
 *   正常档（或反之），比不分档更危险。故拒绝路径显式返回 eInvalid + 置码，
 *   调用方凭 uErrorId 区分"正常档判定"与"拒绝档"，绝不静默输出。
 *
 * 验收向量 (Acceptance) : （fLowLimit=10, fLowWarn=20, fUpWarn=80, fUpLimit=90）
 *   V1 fVal =  5.0 → eLowTripped，uErrorId = 0
 *   V2 fVal = 15.0 → eLowWarn，   uErrorId = 0
 *   V3 fVal = 50.0 → eNormal，    uErrorId = 0
 *   V4 fVal = 85.0 → eUpWarn，    uErrorId = 0
 *   V5 fVal = 95.0 → eUpTripped， uErrorId = 0
 *   V6 阈值组 90/80/20/10（序倒置）→ eInvalid，uErrorId 非 0（拒绝路径验证）
 *
 * 【边界值归属推演表 / Boundary attribution walk-through】
 *   （同一阈值组 10 / 20 / 80 / 90，逐边界值验证闭区间口径 B1）
 *   B1v fVal = 10.0 → eLowTripped（等于低低限，贴线即停机级）
 *   B2v fVal = 20.0 → eLowWarn   （等于低警告限，归更严档）
 *   B3v fVal = 80.0 → eUpWarn    （等于高警告限，归更严档）
 *   B4v fVal = 90.0 → eUpTripped （等于高高限，贴线即停机级）
 *   B5v fVal = 10.000000001      ：高于低低限且容差外 → eLowWarn
 *   B6v fVal = 89.999999999      ：低于高高限且容差外 → eUpWarn
 *
 * 【退化组态语义 / Degenerate configuration semantics】
 *   相邻阈值相等合法，档位按闭区间口径退化收缩：
 *   fLowWarn = fLowLimit = 15 → 低低与低档收缩为同一条线（v <= 15 全判低低）；
 *   fUpWarn = fUpLimit = 85  → 高档与高高档收缩为同一条线（v >= 85 全判高高）；
 *   fLowWarn = fUpWarn = 50  → **正常档退化为空集**：v = 50 被「<= 低警告限」
 *   严档优先拦截判 eLowWarn，v > 50 与 v < 50 两侧分别落入低档 / 高档，
 *   eNormal 无任何取值可达（v1.0.1 终审勘误：原文「仅 v = 50 判正常」与
 *   闭区间归属次序不符，属文档错、代码对）。
 *   退化组态常用于"四线表只用两线"的简化仪表位，属合法工况不置诊断；
 *   序倒置（严格大于）才是组态错误，走 eInvalid 拒绝路径。
 * 故障码表 (Error codes):
 *   16#0001_0214  阈值序非法：要求 fLowLimit <= fLowWarn <= fUpWarn <= fUpLimit，
 *                 相邻阈值倒置（含容差内倒置）即置码，返回 eInvalid，禁止静默分档
 *   【码位终审】原拟 0003_0201 属 DL_Device 段位，且与设备族「非法状态」共用码
 *   （DolMotor / PneumaticCylinder / StarDeltaMotor）语义冲突；本体属 DL_Base，
 *   已顺延至 0001_0214（DL_Base 段 0201~0213 已占用，0214 空闲）。
 * 红线自检 (Redline)    : R1 ✓ 零全局存储 / 零外部变量引用 ｜ R2 ✓ 零物理地址直写
 *                         R3 ✓ 纯 IEC 61131-3 ｜ R4 ✓ 阈值序校验 + 容差判等 + 非法拒绝不静默
 *                         R5 ✓ 全变量与枚举项中英双语同行注释 ｜ R6 ✓ 纯函数无状态（R6 状态机 N/A）
 *                         R7 ✓ 无定时器 / 边沿实例（R7 N/A）
 * 边界契约 (Boundaries):
 *   B1 边界值归属写死：等于阈值归更严档（<= 与 >= 闭区间口径）——
 *      fVal = fLowLimit 判低低档，fVal = fUpLimit 判高高档，fVal = fUpWarn 判高档。
 *      仪表联锁场景"贴线即触发"是安全侧惯例，注释固化不得随实现漂移。
 *   B2 阈值序校验：相邻相等视为合法（档位退化，如 fLowWarn = fUpWarn 时
 *      正常档收缩为一点）；序倒置（严格大于）或容差内倒置判非法，
 *      返回 eInvalid 并置码——分档错误比不分档更危险，禁止静默输出。
 *   B3 纯函数：同输入同输出，无内部状态、无副作用，可安全放进 IF 表达式。
 * 修订历史 (Revision)   :
 *   2026-11-15  v1.0.0  首版落盘（Round 09 · 泳道 A · Level 0 原子族回补）
 *   2026-11-15  v1.0.1  终审修复：故障码 0003_0201 属 DL_Device 段且与设备族
 *                       非法状态码冲突，顺延为 0001_0214；勘误退化组态说明
 *                       （fLowWarn = fUpWarn 时正常档为空集，非"单点"），
 *                       代码行为未改动
 *============================================================================*)
TYPE E_DL_LimitBand :
(
    eLowTripped := 0,  // 低低档：<= 低低限，停机级 / Low-low band, trip level
    eLowWarn    := 1,  // 低档：<= 低警告限 / Low warning band
    eNormal     := 2,  // 正常档 / Normal band
    eUpWarn     := 3,  // 高档：>= 高警告限 / High warning band
    eUpTripped  := 4,  // 高高档：>= 高高限，停机级 / High-high band, trip level
    eInvalid    := 9   // 参数非法兜底档 / Invalid-parameters fallback band
);
END_TYPE

FUNCTION FC_DL_LimitClassify : E_DL_LimitBand   // 返回档位判定结果 / Returns the band judgment
VAR_INPUT
    fVal      : LREAL;                  // 被判定值 [工程单位随应用] / Value to classify [EU by application]
    fLowLimit : LREAL;                  // 低低限（停机级）[工程单位] / Low-low trip limit [EU]
    fLowWarn  : LREAL;                  // 低警告限 [工程单位] / Low warning limit [EU]
    fUpWarn   : LREAL;                  // 高警告限 [工程单位] / High warning limit [EU]
    fUpLimit  : LREAL;                  // 高高限（停机级）[工程单位] / High-high trip limit [EU]
END_VAR
VAR_OUTPUT
    uErrorId  : UDINT;                  // 故障码，0 = 无故障；阈值序非法置码 / Error code, 0 = no error
END_VAR
VAR CONSTANT
    DL_FLOAT_EPS : LREAL := 1.0E-9;     // 判等容差（阈值相邻容差内倒置判非法）/ Equality tolerance for the limit order check
END_VAR

(*------------------------------------------------------------------------------
 * 段 1｜缺省返回：非法兜底档，故障码清零（合法路径再覆盖）
 *      Default return: invalid fallback band, error code cleared first
 *      缺省即拒绝语义：任何未显式分档的退出路径都携带 eInvalid，不误报
 *-----------------------------------------------------------------------------*)
FC_DL_LimitClassify := E_DL_LimitBand.eInvalid;
uErrorId := 16#0000_0000;

(*------------------------------------------------------------------------------
 * 段 2｜阈值序校验（边界 B2）：四阈值须单调不减，倒置或容差内倒置判非法
 *      Limit order check: four limits must be monotonically non-decreasing
 *      容差内倒置（如 fLowWarn 比 fLowLimit 大 1E-12）按倒置处理，
 *      避免浮点噪声吞掉真组态错误
 *-----------------------------------------------------------------------------*)
IF (fLowLimit > fLowWarn + DL_FLOAT_EPS)
    OR (fLowWarn > fUpWarn + DL_FLOAT_EPS)
    OR (fUpWarn > fUpLimit + DL_FLOAT_EPS) THEN
    uErrorId := 16#0001_0214;   // 故障级：阈值序非法 / Fault: invalid limit order
    RETURN;                     // 拒绝路径：保持 eInvalid，禁止静默分档（B2）
END_IF

(*------------------------------------------------------------------------------
 * 段 3｜五档判定主体（边界 B1）：闭区间口径，等于阈值归更严档，
 *      判据全部 ABS 差值与容差比较，禁浮点直接判等
 *      Five-band body with closed-interval attribution, tolerance-based compares
 *-----------------------------------------------------------------------------*)
IF fVal <= fLowLimit THEN
    FC_DL_LimitClassify := E_DL_LimitBand.eLowTripped;      // 贴线即停机级（安全侧，B1）
ELSIF fVal <= fLowWarn THEN
    FC_DL_LimitClassify := E_DL_LimitBand.eLowWarn;         // 低警告档 / Low warning band
ELSIF ABS(fVal - fUpLimit) < DL_FLOAT_EPS THEN
    FC_DL_LimitClassify := E_DL_LimitBand.eUpTripped;       // 等于高高限归更严档（容差判等）
ELSIF fVal >= fUpLimit THEN
    FC_DL_LimitClassify := E_DL_LimitBand.eUpTripped;       // 超高高限 / Above high-high
ELSIF ABS(fVal - fUpWarn) < DL_FLOAT_EPS THEN
    FC_DL_LimitClassify := E_DL_LimitBand.eUpWarn;          // 等于高警告限归更严档（容差判等）
ELSIF fVal >= fUpWarn THEN
    FC_DL_LimitClassify := E_DL_LimitBand.eUpWarn;          // 高警告档 / High warning band
ELSE
    FC_DL_LimitClassify := E_DL_LimitBand.eNormal;          // 正常档 / Normal band
END_IF
(* 到此全部分档路径已覆盖：低低 / 低 / 高高 / 高 / 正常五档互斥完备，
   容差分支仅在上边界两侧生效，低侧由 <= 闭区间天然覆盖等值归属 *)
END_FUNCTION

(* ---- FC_DL_WordBitPack.st ---- *)
(*==============================================================================
 * 组件名称 (Component)  : FC_DL_WordBitPack
 * 所属子库 (Sublibrary) : DL_Base
 * 当前版本 (Version)    : 1.0.1
 * 分类     (Category)   : 位逻辑纯函数（Function · Bit Logic）
 * 兼容性   (Platform)   : CODESYS 3.5 / TwinCAT 3 / 汇川 InoProShop / Machine Expert
 *                         仅依赖 Standard.library（SHL / SHR / AND / OR / NOT），
 *                         零厂商方言
 * 功能简介 (Function)   : 按位偏移 + 位宽参数把字段值合入目标字（打包），同拍
 *                         经输出引脚回读该位段旧值（解包），一个函数完成
 *                         「读-改-写」原子语义：uExtracted 给出改动前的位段
 *                         内容，返回值给出改动后的整字。字段值右对齐，超出
 *                         位宽的高位被掩码忽略。偏移+宽度越界或宽度为 0 时
 *                         拒绝执行：返回原字不动、uExtracted 返回 0、置故障码
 *                         （禁止半写，防位段被撕裂）。纯函数：无状态、无副作用。
 *                         与已入库 FC_DL_PackBitsToWord（16 点 BOOL 打包整字）、
 *                         FB_DL_UnpackWordToBits（整字展开 16 点）职责分离——
 *                         本块是任意位段（偏移/宽度参数化）的打包解包原子。
 * 开源溯源 (Origin)     : 原创实现（参考 LGF 库 Bit Logic 位逻辑分类的功能域
 *                         与参数域，来源标签 lgf-bitlogic），读-改-写掩码法为
 *                         公开经典位运算手法，仅借分类/参数域/命名，clean-room
 *                         实现，未复制任何厂商私有库源码，不构成衍生作品。
 * 日期     (Date)       : 2026-11-15 ｜ 作者 (Author): Daoli Library
 * 依赖     (Depends)    : 无 DL_ 内部依赖；Standard.library: SHL / SHR / AND / OR / NOT
 *
 *------------------------------------------------------------------------------
 * 【引脚契约 / Pin contract】
 *   输入 uTarget    : WORD  — 目标载体字（旧内容），打包基址；
 *   输入 uField     : WORD  — 待合入字段值（右对齐，超出位宽的高位被忽略）；
 *   输入 nOffset    : USINT — 位段起始偏移 [bit]，合法域 0~15；
 *   输入 nWidth     : USINT — 位段宽度 [bit]，合法域 1~16；
 *   输出 uExtracted : WORD  — 该位段的旧值（右对齐回读，即解包结果）；
 *   输出 uErrorId   : UDINT — 故障码，0 = 无故障；16#0001_0108 = 位段越界拒绝；
 *   返回值          : WORD  — 合成后的字（拒绝路径返回原字不动）。
 *
 * 【边界防错清单 / Boundary guard list】
 *   B1 nWidth = 0 或 nWidth > 16 或 nOffset >= 16 或 nOffset + nWidth > 16 →
 *      置故障，返回原字不动、uExtracted 返回 0（禁止半写：宁可整拍不动，
 *      绝不撕裂位段）。四项判据缺一不可：nWidth / nOffset 引脚类型为 USINT
 *      （域 0~255），若只判 nOffset + nWidth > 16，则 15 + 250 = 265 在 USINT
 *      域内回绕成 9 从而漏判，随后 SHL 位移 250 位落入平台未定义行为
 *      （v1.0.1 终审补齐，原 v1.0.0 只有两项判据）。
 *   B2 掩码构造：宽度 16 时左移 16 位行为按「满宽度掩码显式分支」处理，
 *      不依赖平台移位语义（部分平台 SHL(x,16) 结果为 0 或回绕，口径不一）；
 *   B3 字段值合入前先按位段宽度掩码截断（高位越宽忽略），再左移对齐；
 *   B4 纯函数无状态，同输入同输出；拒绝路径输入输出零修改；
 *   B5 逐项判界后 nOffset <= 15 且 nWidth <= 16，加法上界 31 不越 USINT 域，
 *      全部移位计数值严格小于 16（平台无关）。
 *
 * 【原子语义声明 / Atomic semantics】
 *   「读-改-写」原子指单次调用内完成三步：读（uExtracted 回读旧位段）、
 *   改（掩码清旧段）、写（新字段值入段）；调用方在同一表达式中同时取得
 *   改前值与改后值，无需两次调用，避免了两次调用之间字段值被外部修改的
 *   时序缝隙。注意：原子性限于本函数单次调用内部，跨多个调用方的整字
 *   互斥仍需上层仲裁（本函数不持锁、不触碰任何共享存储）。
 *
 * 【调用示例 / Call example】
 *   「把模式号 3 写入状态字的 bit4~bit7，同时留档旧模式」
 *   wOldMode := FC_DL_WordBitPack(uTarget := wStatus, uField := 3,
 *                                 nOffset := 4, nWidth := 4,
 *                                 uExtracted => wOldMode, uErrorId => uErr);
 *
 * 【平台移植注意 / Porting notes】
 *   各平台 SHL/SHR 对移位计数 ≥ 数据宽度的行为定义不一（结果 0 / 回绕 /
 *   未定义），本函数通过边界 B1（越界拒绝）与 B2（满宽度显式分支）从设计上
 *   规避了该平台差异，全部移位计数值均严格小于 16，不触发任何方言行为。
 *
 * 【同族职责分离 / Family separation】
 *   FC_DL_PackBitsToWord：16 点 BOOL → 整字（固定全字打包，无偏移参数）；
 *   FB_DL_UnpackWordToBits：整字 → 16 点 BOOL（固定全字解包）；
 *   本函数：任意位段（偏移/宽度参数化）打包 + 解包回读，三者正交不互调。
 *
 * 红线自检 (Redline)    : R1 零全局变量表/外部变量引用 ✓ ｜ R2 零物理 IO 地址 ✓
 *                         R3 纯 IEC 61131-3 标准位运算 ✓ ｜ R4 越界拒绝禁半写/
 *                           出口唯一/无除法/循环界常量无死锁 ✓
 *                         R5 全变量中英双语同行注释 ✓ ｜ R6 N/A（纯函数无状态机）
 *                         R7 N/A（无定时器/边沿实例）｜ R8 位宽/偏移/掩码全常量化 ✓
 * 验收向量 (Acceptance) :
 *   V1  uTarget=16#0000, uField=16#3,  nOffset=4,  nWidth=4
 *       → 返回 16#0030, uExtracted = 16#0000, uErrorId = 0
 *   V2  uTarget=16#00FF, uField=16#0,  nOffset=0,  nWidth=8
 *       → 返回 16#0000, uExtracted = 16#00FF, uErrorId = 0
 *   V3  uTarget=16#0000, uField=16#F,  nOffset=12, nWidth=4
 *       → 返回 16#F000, uExtracted = 16#0000, uErrorId = 0
 *   V4  uTarget=16#1234, uField=16#A,  nOffset=4,  nWidth=4
 *       → 返回 16#12A4, uExtracted = 16#0003, uErrorId = 0
 *   V5  uTarget=16#1234, uField=16#AA, nOffset=4,  nWidth=5
 *       → 返回 16#12A4, uExtracted = 16#0003, uErrorId = 0
 *       【验算注记 / Verification note】ROUND_PLAN_R9 §9 V5 表原载期望返回
 *       16#1264；按「右对齐 + 超宽高位忽略」语义逐位验算：
 *         掩码 = 5 个 1 左移 4 位           = 16#01F0
 *         uField 16#AA 截低 5 位（16#AA AND 16#1F）= 16#0A
 *         字段左移 4 位                     = 16#00A0
 *         载体清段 16#1234 AND NOT 16#01F0  = 16#1204
 *         合成 16#1204 OR 16#00A0           = 16#12A4
 *       【R9 终审裁定 / Final ruling】总监逐位独立复核，结果 16#12A4：位 4~8
 *       由 0_1010 覆盖后为 0001_0010_1010_0100。16#1264 的位 4~8 = 0_0110
 *       （字段值 6），与本组入参 16#AA、宽度 5、偏移 4 无任何推导路径，
 *       判定为**计划向量笔误**：代码对、向量错。已同步勘误 ROUND_PLAN_R9.md
 *       §9 V5 表（16#1264 → 16#12A4 并附勘误脚注），保留 R8「公式对、
 *       向量错」口径的勘误留痕；本组件实现不做改动。
 *   V6  uTarget=16#1234, uField=16#1,  nOffset=15, nWidth=2
 *       → 返回 16#1234（原字不动）, uExtracted = 16#0000,
 *         uErrorId = 16#0001_0108（偏移+宽度越界拒绝）
 *   V7  uTarget=16#1234, uField=16#1,  nOffset=15, nWidth=250（v1.0.1 新增）
 *       → 返回 16#1234（原字不动）, uExtracted = 16#0000,
 *         uErrorId = 16#0001_0108（宽度单项越界拒绝；若只判「偏移+宽度>16」，
 *         15+250 在 USINT 域回绕为 9 会漏判，故宽度 / 偏移各自设界）
 *
 * 【故障码表 / Error code table】
 *   16#0001_0108  位段越界拒绝：nWidth = 0 / nWidth > 16 / nOffset >= 16 /
 *                 nOffset + nWidth > 16，返回原字不动、uExtracted = 0，
 *                 瞬时码每次调用重算（0108 空闲，0101~0107 已被计数/步进/
 *                 BCD 族登记，0109 已被 MonthWindowCheck 登记，010A 起空闲）。
 *
 * 【实现选择 / Implementation choice】
 *   两掩码法：段掩码 uMask = width 个 1 左移 offset（清旧段 + 提旧值共用），
 *   字段掩码 uFieldMask = SHR(uMask, nOffset)（截断超宽高位）；合成式
 *   (uTarget AND NOT uMask) OR SHL(uField AND uFieldMask, nOffset)，三个
 *   中间量全部显式命名，无嵌套魔法表达式；满宽度（width = 16）走显式分支
 *   直接赋 16#FFFF，规避平台移位语义差异（边界 B2）。
 *
 * 【逐步验算表 / Step-by-step walkthrough（供终审逐组代回验算）】
 *   V1 掩码 16#00F0；uExtracted = 0；清段 0；合段 3<<4 = 16#0030 ✓
 *   V2 掩码 16#00FF；uExtracted = 16#00FF；清段后 0；合段 0 → 16#0000 ✓
 *   V3 掩码 16#F000；uExtracted = 0；合段 16#F<<12 = 16#F000 ✓
 *   V4 掩码 16#00F0；uExtracted = (16#34 AND 16#F0)>>4 = 3；
 *      清段 16#1204；合段 16#A<<4 = 16#A0 → 16#12A4 ✓
 *   V5 掩码 16#01F0；uExtracted = (16#34 AND 16#F0)>>4 = 3；
 *      字段截断 16#AA AND SHR(16#01F0,4) = 16#AA AND 16#1F = 16#0A；
 *      清段 16#1204；合段 16#0A<<4 = 16#A0 → 16#12A4（差异注记见上）✓
 *   V6 15 + 2 = 17 > 16 → 拒绝：原字 16#1234 原样返回、uExtracted = 0、
 *      置 0001_0108 ✓
 *
 * 修订历史 (Revision)   :
 *   2026-11-15  v1.0.0  首版落盘（Round 09 · 泳道 A · LGF Bit Logic 组）
 *   2026-11-15  v1.0.1  终审修复：参数防御补「nWidth > 16」「nOffset >= 16」
 *                       两项单项判界（原实现只判 nOffset + nWidth > 16，USINT
 *                       域 15 + 250 回绕为 9 可绕过校验并触发平台未定义移位）；
 *                       同步落定 V5 向量裁定（计划表 16#1264 → 代码实测语义
 *                       16#12A4，计划文件已勘误）
 *============================================================================*)
FUNCTION FC_DL_WordBitPack : WORD          // 返回合成后的字 / Returns the assembled word
VAR_INPUT
    uTarget  : WORD;                       // 目标载体字（旧内容）/ Target carrier word (previous content)
    uField   : WORD;                       // 待合入字段值，右对齐，超宽高位被忽略 / Field value to merge, right-aligned, bits above width ignored
    nOffset  : USINT;                      // 位段起始偏移 [bit]，合法域 0~15 / Field start offset [bit], legal range 0~15
    nWidth   : USINT;                      // 位段宽度 [bit]，合法域 1~16 / Field width [bit], legal range 1~16
END_VAR
VAR_OUTPUT
    uExtracted : WORD;                     // 该位段旧值，右对齐回读（解包结果）/ Previous field value, right-aligned (unpack result)
    uErrorId   : UDINT;                    // 故障码，0 = 无故障，0001_0108 = 越界拒绝 / Error code, 0 = none, 0001_0108 = out-of-range rejected
END_VAR
VAR
    uMask      : WORD;                     // 位段掩码：width 个 1 左移 offset / Field mask: width ones shifted left by offset
    uMaskInv   : WORD;                     // 掩码反相：清旧段用 / Inverted mask for clearing the old field
    uFieldMask : WORD;                     // 字段掩码：段掩码右对齐，截超宽高位 / Field-side mask, right-aligned, truncates oversized bits
    uFieldTrim : WORD;                     // 截断后的字段值（右对齐）/ Trimmed field value (right-aligned)
    uFieldAlgn : WORD;                     // 对齐后的字段值（左移 offset）/ Aligned field value (shifted left by offset)
    uBase      : WORD;                     // 清段后的载体字 / Carrier word with the old field cleared
    bValid     : BOOL;                     // 参数合法标志（拒绝路径闸门）/ Parameter validity flag (rejection-path gate)
END_VAR
VAR CONSTANT
    DL_WORD_BITS : USINT := 16;            // WORD 位宽 [bit] / Width of a WORD [bit]
    DL_WORD_FULL : WORD  := 16#FFFF;       // 满字掩码（宽度 16 显式分支用）/ Full-word mask for the explicit width-16 branch
    DL_BIT_ONE   : WORD  := 16#0001;       // 单位种子（掩码构造显式 WORD 化，防字面量平台默认类型差异）/ One-bit seed, explicit WORD typing to avoid platform literal defaults
    DL_BIT_ERR_RNG: UDINT := 16#0001_0108; // 位段越界拒绝故障码 / Error code for out-of-range rejection
END_VAR

(*------------------------------------------------------------------------------
 * 段 1｜安全预置（P-01 范式）：拒绝路径返回原字、uExtracted 返回 0
 *      Safe preset: rejection paths return the original word, uExtracted = 0
 *-----------------------------------------------------------------------------*)
uErrorId     := 16#0000_0000;              // 故障码预清零，正常路径末尾保持 0 / Error code preset to zero, stays 0 on the normal path
uExtracted   := 16#0000;                   // 解包结果预清零，合法路径段 3 回读覆盖 / Unpack result preset to zero, overwritten by stage 3 on legal paths
bValid       := TRUE;                      // 参数合法性预置为通过（Validity preset to pass）

(*------------------------------------------------------------------------------
 * 段 2｜参数防御（边界 B1）：宽度 0 / 宽度 > 16 / 偏移 >= 16 / 偏移+宽度 > 16
 *      任一命中即整体拒绝，禁半写
 *      Parameter guard (B1): zero width, width above 16, offset at or above 16,
 *      or offset plus width above 16 rejects the whole call
 *      单项判界先于求和判界：USINT 域内 15 + 250 = 265 会回绕成 9，
 *      只判求和会漏判并让 SHL 移位 250 位落入平台未定义行为（v1.0.1 补齐）
 *      Single checks precede the sum check because the USINT sum wraps
 *-----------------------------------------------------------------------------*)
IF (nWidth = 0) OR (nWidth > DL_WORD_BITS) OR (nOffset >= DL_WORD_BITS) OR
   (nOffset + nWidth > DL_WORD_BITS) THEN
    bValid   := FALSE;                     // 参数非法，置拒绝闸门 / Invalid parameters, close the rejection gate
    uErrorId := DL_BIT_ERR_RNG;            // 置位段越界拒绝故障码 / Raise out-of-range rejection code
END_IF

IF bValid THEN
    (*--------------------------------------------------------------------------
     * 段 3｜解包回读（读）：旧位段右对齐提取，同拍返回给调用方留档
     *      Unpack read-back (read): old field extracted right-aligned
     *-------------------------------------------------------------------------*)
    IF nWidth = DL_WORD_BITS THEN
        uMask := DL_WORD_FULL;             // 满宽度显式分支：直接全字掩码 / Explicit width-16 branch: full-word mask directly
    ELSE
        uMask := SHL(SHL(DL_BIT_ONE, nWidth) - 1, nOffset); // width 个 1 左移 offset（种子显式 WORD 化）/ width ones shifted left by offset (explicit WORD seed)
    END_IF
    uMaskInv := NOT uMask;                 // 掩码反相，清旧段用 / Invert mask for clearing the old field
    uExtracted := SHR(uTarget AND uMask, nOffset); // 旧位段右对齐回读 / Read back old field, right-aligned

    (*--------------------------------------------------------------------------
     * 段 4｜打包合成（改 + 写）：清旧段 → 字段截断 → 对齐 → 按位或
     *      Pack and merge (modify + write): clear, trim, align, merge
     *   单步数据流：
     *     uTarget AND uMaskInv ──► uBase（旧段清零的载体）
     *     uFieldMask = SHR(uMask, nOffset)（段掩码右对齐）
     *     uField AND uFieldMask ──► uFieldTrim（超宽高位忽略）
     *     uFieldTrim SHL nOffset ──► uFieldAlgn（对齐到目标位段）
     *     uBase OR uFieldAlgn ──► 返回值（合成后的字）
     *-------------------------------------------------------------------------*)
    uBase      := uTarget AND uMaskInv;    // 载体字清旧段（载体 cleared of old field）
    uFieldMask := SHR(uMask, nOffset);     // 段掩码右对齐（mask aligned to field side）
    uFieldTrim := uField AND uFieldMask;   // 字段截断，超宽高位忽略（trim oversized bits）
    uFieldAlgn := SHL(uFieldTrim, nOffset); // 字段对齐到目标位段（align field to target bits）
    FC_DL_WordBitPack := uBase OR uFieldAlgn; // 读-改-写合成出口 / Read-modify-write merge exit
ELSE
    FC_DL_WordBitPack := uTarget;          // 拒绝路径：原字原样返回，禁半写 / Rejection path: return the original word untouched
END_IF

(*------------------------------------------------------------------------------
 * 段 5｜出口一致性（边界 B4）：唯一出口，拒绝与合法路径互不残留
 *      Exit consistency (B4): single exit, no cross-path residue
 *-----------------------------------------------------------------------------*)
(* 拒绝路径时 uExtracted 保持段 1 预置的 0，合法路径为段 3 回读旧值：
   两条路径的 uExtracted 语义均在头注释契约中写死，无隐式行为 *)
END_FUNCTION
